FUNCTION "HMI COMMS" : VOID
TITLE =HMI Communications
//OMRON NS12  on DB12
NAME : HMI_COMM
VERSION : 0.1


VAR_TEMP
  UPDATE_PULSE_0 : BOOL ;
  UPDATE_PULSE_1 : BOOL ;
  UPDATE_PULSE_2 : BOOL ;
  UPDATE_PULSE_3 : BOOL ;
  UPDATE_PULSE_4 : BOOL ;
  UPDATE_PULSE_5 : BOOL ;
  UPDATE_PULSE_6 : BOOL ;
  UPDATE_1 : BOOL ;
  UPDATE_2 : BOOL ;
  UPDATE_3 : BOOL ;
  UPDATE_4 : BOOL ;
  UPDATE_5 : BOOL ;
  UPDATE_6 : BOOL ;
  UPDATE_7 : BOOL ;
  UPDATE_8 : BOOL ;
  UPDATE_9 : BOOL ;
  UPDATE_10 : BOOL ;
  UPDATE_11 : BOOL ;
  UPDATE_12 : BOOL ;
  UPDATE_13 : BOOL ;
  TEMP1 : BOOL ;
  TEST : BOOL ;
  CONVEYOR_0_COLOR : BYTE ;
  ELEVATOR_COLOR : BYTE ;
  CONVEYOR_1_COLOR : BYTE ;
  CONVEYOR_2_COLOR : BYTE ;
  CONVEYOR_3_COLOR : BYTE ;
  CONVEYOR_4_COLOR : BYTE ;
  CONVEYOR_5_COLOR : BYTE ;
  CONVEYOR_6_COLOR : BYTE ;
  CONVEYOR_7_COLOR : BYTE ;
  CONVEYOR_8_COLOR : BYTE ;
  CONVEYOR_9_COLOR : BYTE ;
  PUSHER_2_COLOR : BOOL ;
  CONVEYOR_11_COLOR : BYTE ;
  CONVEYOR_12_COLOR : BYTE ;
  CONVEYOR_13_COLOR : BYTE ;
  CONVEYOR_21_COLOR : BYTE ;
  CONVEYOR_22_COLOR : BYTE ;
  CONVEYOR_23_COLOR : BYTE ;
  CONVEYOR_10_COLOR : BYTE ;
  NEW_ORDER_COLOR : BYTE ;
END_VAR
BEGIN
NETWORK
TITLE =HMI - UpDate Timing
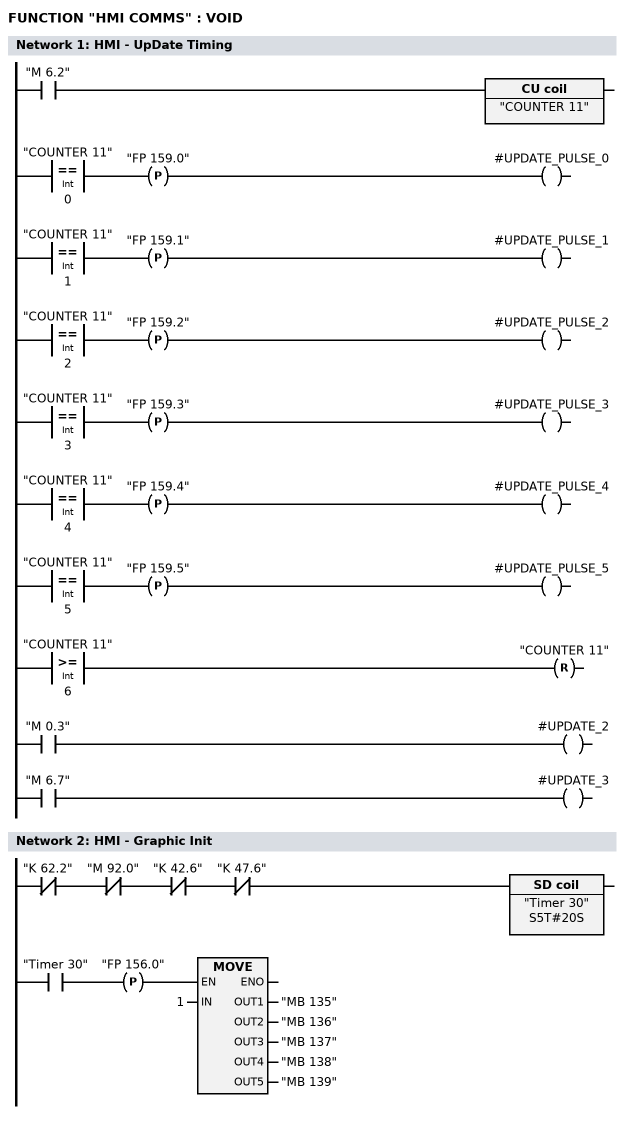

      A     "M 6.2";
      CU    "COUNTER 11";
//;
      A(    ;
      L     "COUNTER 11";
      L     0;
      ==I   ;
      )     ;
      FP    "FP 159.0";
      =     #UPDATE_PULSE_0;
//;
      A(    ;
      L     "COUNTER 11";
      L     1;
      ==I   ;
      )     ;
      FP    "FP 159.1";
      =     #UPDATE_PULSE_1;
//;
      A(    ;
      L     "COUNTER 11";
      L     2;
      ==I   ;
      )     ;
      FP    "FP 159.2";
      =     #UPDATE_PULSE_2;
//;
      A(    ;
      L     "COUNTER 11";
      L     3;
      ==I   ;
      )     ;
      FP    "FP 159.3";
      =     #UPDATE_PULSE_3;
//;
      A(    ;
      L     "COUNTER 11";
      L     4;
      ==I   ;
      )     ;
      FP    "FP 159.4";
      =     #UPDATE_PULSE_4;
//;
      A(    ;
      L     "COUNTER 11";
      L     5;
      ==I   ;
      )     ;
      FP    "FP 159.5";
      =     #UPDATE_PULSE_5;
//;
      A(    ;
      L     "COUNTER 11";
      L     6;
      >=I   ;
      )     ;
      R     "COUNTER 11";
//;;
      A     "M 0.3";
      =     #UPDATE_2;
//;
      A     "M 6.7";
      =     #UPDATE_3;
NETWORK
TITLE =HMI - Graphic Init

      AN    "K 62.2";
      AN    "M 92.0";
      AN    "K 42.6";
      AN    "K 47.6";
      L     S5T#20S;
      SD    "Timer 30";
//;
      A     "Timer 30";
      FP    "FP 156.0";
      JNB   K622;
      L     1;
      T     "MB 135";
      T     "MB 136";
      T     "MB 137";
      T     "MB 138";
      T     "MB 139";

K622: NOP   0;
NETWORK
TITLE =HMI - Doors Monitor

      ON    "E 4.6";
      ON    "E 9.0";
      ON    "E 12.5";
      O     #UPDATE_PULSE_0;
      JNB   DOOR;
      AN    "E 4.6";
      =     "HMI_DB".ELEVATOR_DOOR_STATUS;
//;
      AN    "E 9.0";
      =     "HMI_DB".FLIPPER_DOOR_STATUS;
//;
      AN    "E 12.5";
      =     "HMI_DB".LOADER_DOOR_STATUS;

DOOR: NOP   0;
NETWORK
TITLE =HMI - E-Stop Monitor

      O     "M 1.0";
      O     "M 1.1";
      O     "M 1.2";
      O     "M 1.3";
      O     #UPDATE_PULSE_1;
      JNB   ESTP;
      A     "M 1.0";
      =     "HMI_DB".E_STOP_CONSOLE_STATUS;
//;
      A     "M 1.1";
      =     "HMI_DB".E_STOP_LOADER_STATUS;
//;
      A     "M 1.2";
      =     "HMI_DB".E_STOP_ELEVATOR_STATUS;
//;
      A     "M 1.3";
      =     "HMI_DB".E_STOP_FLIPPER_STATUS;

ESTP: NOP   0;
NETWORK
TITLE =HMI - Motors Fault Status

      A(    ;
      L     "MW 2";
      L     0;
      <>I   ;
      O     ;
      L     "MB 4";
      L     0;
      <>I   ;
      )     ;
      O     "M 7.0";
      O     "M 7.1";
      O     "M 7.2";
      O     #UPDATE_PULSE_2;
      JNB   MTRF;
      A     "M 2.0";
      =     "HMI_DB".CONVEYOR_0_MOTOR_STATUS;
//;
      A     "M 2.1";
      =     "HMI_DB".PUSHER_0_MOTOR_STATUS;
//;
      A     "M 2.2";
      =     "HMI_DB".ELEVATOR_MOTOR_STATUS;
//;
      A     "M 2.3";
      =     "HMI_DB".PUSHER_1_MOTOR_STATUS;
//;
      A     "M 2.4";
      =     "HMI_DB".CONVEYOR_1_MOTOR_STATUS;
//;
      A     "M 2.5";
      =     "HMI_DB".CONVEYOR_2B_MOTOR_STATUS;
//;
      A     "M 2.6";
      =     "HMI_DB".CONVEYOR_2R_MOTOR_STATUS;
//;
      A     "M 2.7";
      =     "HMI_DB".CONVEYOR_3_MOTOR_STATUS;
//;
      A     "M 3.0";
      =     "HMI_DB".CONVEYOR_4_MOTOR_STATUS;
//;
      A     "M 3.1";
      =     "HMI_DB".CONVEYOR_5_MOTOR_STATUS;
//;
      A     "M 3.2";
      =     "HMI_DB".CONVEYOR_6_MOTOR_STATUS;
//;
      A     "M 3.3";
      =     "HMI_DB".CONVEYOR_7_MOTOR_STATUS;
//;
      A     "M 3.4";
      =     "HMI_DB".FLIPPER_MOTOR_STATUS;
//;
      A     "M 3.5";
      =     "HMI_DB".CONVEYOR_8_MOTOR_STATUS;
//;
      A     "M 3.6";
      =     "HMI_DB".TURNTABLE_MOTOR_STATUS;
//;
      A     "M 3.7";
      =     "HMI_DB".CONVEYOR_9_MOTOR_STATUS;
//;
      A     "M 4.0";
      =     "HMI_DB".PUSHER_2_MOTOR_STATUS;
//;
      A     "M 4.1";
      =     "HMI_DB".CONVEYOR_10_MOTOR_STATUS;
//;
      A     "M 4.2";
      =     "HMI_DB".CONVEYOR_11_MOTOR_STATUS;
//;
      A     "M 4.3";
      =     "HMI_DB".CONVEYOR_12_MOTOR_STATUS;
//;
      A     "M 4.4";
      =     "HMI_DB".CONVEYOR_13_MOTOR_STATUS;
//;
      A     "M 4.5";
      =     "HMI_DB".CONVEYOR_21_MOTOR_STATUS;
//;
      A     "M 4.6";
      =     "HMI_DB".CONVEYOR_22_MOTOR_STATUS;
//;
      A     "M 4.7";
      =     "HMI_DB".CONVEYOR_23_MOTOR_STATUS;
//;
      A     "M 7.0";
      =     "HMI_DB".LOADER_LIFT_MOTOR_STATUS;
//;
      A     "M 7.1";
      =     "HMI_DB".LOADER_FING_MOTOR_STATUS;
//;
      A     "M 7.2";
      =     "HMI_DB".LOADER_BELT_MOTOR_STATUS;

MTRF: NOP   0;
NETWORK
TITLE =HMI Light Barriers Status - Conveyors 1, 2, 3 LBs

      A(    ;
      L     IW     5;
      L     "HMI_UPDATE".HMI_GRAPHIC_TOTAL_1;
      <>I   ;
      O     #UPDATE_PULSE_3;
      )     ;
      JNB   LBS1;
      A     "B 5.4";
      =     "HMI_DB".LIGHT_BARRIER_1_STATUS;
//;
      A     "B 5.5";
      =     "HMI_DB".LIGHT_BARRIER_2_STATUS;
//;
      A     "B 6.0";
      =     "HMI_DB".LIGHT_BARRIER_3_STATUS;
//;
      A     "B 6.1";
      =     "HMI_DB".LIGHT_BARRIER_4_STATUS;
//;
      A     "B 6.2";
      =     "HMI_DB".LIGHT_BARRIER_5_STATUS;
//;
      A     "B 6.4";
      =     "HMI_DB".LIGHT_BARRIER_6_STATUS;
//;
      A     "B 5.2";
      =     "HMI_DB".LIGHT_BARRIER_B_STATUS;
//;
      A     "B 5.1";
      =     "HMI_DB".LIGHT_BARRIER_A_STATUS;
//;
      L     IW     5;
      T     "HMI_UPDATE".HMI_GRAPHIC_TOTAL_1;

LBS1: NOP   0;
NETWORK
TITLE =HMI Light Barriers Status - Conveyors 4, 5, 6, 7, 8, 9 LBs

      A(    ;
      L     IW     6;
      L     "HMI_UPDATE".HMI_GRAPHIC_TOTAL_2;
      <>I   ;
      O     #UPDATE_PULSE_4;
      )     ;
      O     "B 8.2";
      JNB   LBS2;
      A     "B 6.7";
      =     "HMI_DB".LIGHT_BARRIER_7_STATUS;
//;
      A     "B 7.0";
      =     "HMI_DB".LIGHT_BARRIER_8_STATUS;
//;
      A     "B 7.1";
      =     "HMI_DB".LIGHT_BARRIER_9_STATUS;
//;
      A     "B 7.2";
      =     "HMI_DB".LIGHT_BARRIER_10_STATUS;
//;
      A     "B 7.3";
      =     "HMI_DB".LIGHT_BARRIER_11_STATUS;
//;
      A     "B 7.4";
      =     "HMI_DB".LIGHT_BARRIER_12_STATUS;
//;
      A     "B 8.2";
      =     "HMI_DB".LIGHT_BARRIER_13_STATUS;
//;
      L     IW     6;
      T     "HMI_UPDATE".HMI_GRAPHIC_TOTAL_2;

LBS2: NOP   0;
NETWORK
TITLE =HMI Light Barriers Status - Conveyors 10, 11, 12, 13, 21, 22, 23

      A(    ;
      L     IW     9;
      L     IW    12;
      +I    ;
      L     IB    15;
      +I    ;
      L     "HMI_UPDATE".HMI_FEED_GRAPHIC;
      <>I   ;
      O     #UPDATE_PULSE_5;
      )     ;
      JNB   LBS3;
      A     "B 9.6";
      =     "HMI_DB".LIGHT_BARRIER_14_STATUS;
//;
      A     "B 9.7";
      =     "HMI_DB".LIGHT_BARRIER_15_STATUS;
//;
      A     "B 10.3";
      =     "HMI_DB".LIGHT_BARRIER_16_STATUS;
//;
      A     "B 10.4";
      =     "HMI_DB".LIGHT_BARRIER_17_STATUS;
//;
      A     "B 10.5";
      =     "HMI_DB".LIGHT_BARRIER_18_STATUS;
//;
      A     "B 10.6";
      =     "HMI_DB".LIGHT_BARRIER_19_STATUS;
//;
      A     "B 10.7";
      =     "HMI_DB".LIGHT_BARRIER_20_STATUS;
//;
      A     "B 11.0";
      =     "HMI_DB".LIGHT_BARRIER_21_STATUS;
//;
      A     "B 11.1";
      =     "HMI_DB".LIGHT_BARRIER_22_STATUS;
//;
      A     "B 11.2";
      =     "HMI_DB".LIGHT_BARRIER_23_STATUS;
//;
      A     "B 12.3";
      =     "HMI_DB".LIGHT_BARRIER_24_STATUS;
//;
      A     "B 13.0";
      =     "HMI_DB".LIGHT_BARRIER_25_STATUS;
//;
      A     "B 15.4";
      =     "HMI_DB".LIGHT_BARRIER_26_STATUS;
//;
      A     "B 15.5";
      =     "HMI_DB".LIGHT_BARRIER_27_STATUS;
//;
      A     "B 15.6";
      =     "HMI_DB".LIGHT_BARRIER_28_STATUS;
//;
      A     "B 15.7";
      =     "HMI_DB".LIGHT_BARRIER_29_STATUS;
//;
      L     IW     9;
      L     IW    12;
      +I    ;
      L     IB    15;
      +I    ;
      T     "HMI_UPDATE".HMI_FEED_GRAPHIC;

LBS3: NOP   0;
NETWORK
TITLE =HMI Light Barriers Status - Conveyors 0 LBs

      A(    ;
      L     QB    62;
      L     "HMI_UPDATE".HMI_MOTOR_TOTAL_1;
      <>I   ;
      O     #UPDATE_PULSE_0;
      )     ;
      O     "B 8.2";
      JNB   LBS4;
      A     "E 34.7";
      =     "HMI_DB".PACKETIZER_GATE_STATUS;
//;
      A     "B 35.2";
      =     "HMI_DB".LIGHT_BARRIER_30_STATUS;
//;
      A     "B 35.3";
      =     "HMI_DB".LIGHT_BARRIER_31_STATUS;
//;
      A     "B 35.4";
      =     "HMI_DB".LIGHT_BARRIER_32_STATUS;
//;
      L     QB    62;
      T     "HMI_UPDATE".HMI_MOTOR_TOTAL_1;

LBS4: NOP   0;
NETWORK
TITLE =HMI Prox Sensors Status - Elevator - Proxs

      A(    ;
      L     IB     4;
      L     "HMI_UPDATE".HMI_ELEVATOR_PROXS;
      <>I   ;
      O     #UPDATE_PULSE_1;
      )     ;
      JNB   PRX1;
      AN    "P 4.0";
      =     "HMI_DB".PROX_1_STATUS;
//;
      AN    "P 4.1";
      =     "HMI_DB".PROX_2_STATUS;
//;
      AN    "P 4.2";
      =     "HMI_DB".PROX_3_STATUS;
//;
      AN    "P 4.3";
      =     "HMI_DB".PROX_4_STATUS;
//;
      AN    "P 4.4";
      =     "HMI_DB".PROX_5_STATUS;
//;
      AN    "P 4.5";
      =     "HMI_DB".PROX_6_STATUS;
//;
      L     IB     4;
      T     "HMI_UPDATE".HMI_ELEVATOR_PROXS;

PRX1: NOP   0;
NETWORK
TITLE =HMI Prox Sensors Status - Flipper / TurnTable - Proxs

      A(    ;
      L     IW     8;
      L     "HMI_UPDATE".HMI_FLIPPER_PROXS;
      <>I   ;
      O     #UPDATE_PULSE_2;
      )     ;
      JNB   PRX2;
      AN    "P 8.0";
      =     "HMI_DB".PROX_8_STATUS;
//;
      AN    "P 8.1";
      =     "HMI_DB".PROX_7_STATUS;
//;
      AN    "P 8.5";
      =     "HMI_DB".PROX_9_STATUS;
//;
      AN    "P 8.6";
      =     "HMI_DB".PROX_10_STATUS;
//;
      AN    "P 9.2";
      =     "HMI_DB".PROX_11_STATUS;
//;
      AN    "P 9.3";
      =     "HMI_DB".PROX_12_STATUS;
//;
      L     IW     8;
      T     "HMI_UPDATE".HMI_FLIPPER_PROXS;

PRX2: NOP   0;
NETWORK
TITLE =HMI Prox Sensors Status - Pusher 2 / Pivot 10 - Proxs

      A(    ;
      L     IB    10;
      L     IB    15;
      +I    ;
      L     "HMI_UPDATE".HMI_PUSHER_PROXS;
      <>I   ;
      O     #UPDATE_PULSE_3;
      )     ;
      JNB   PRX3;
      AN    "P 10.0";
      =     "HMI_DB".PROX_13_STATUS;
//;
      AN    "P 10.1";
      =     "HMI_DB".PROX_14_STATUS;
//;
      A     "P 15.0";
      =     "HMI_DB".PROX_15_STATUS;
//;
      A     "P 15.1";
      =     "HMI_DB".PROX_16_STATUS;
//;
      L     IB    10;
      L     IB    15;
      +I    ;
      T     "HMI_UPDATE".HMI_PUSHER_PROXS;

PRX3: NOP   0;
NETWORK
TITLE =HMI Prox Sensors Status - Feeder - Proxs

      A(    ;
      L     IW    11;
      L     IB    13;
      +I    ;
      L     "HMI_UPDATE".HMI_FEEDER_PROXS;
      <>I   ;
      O     #UPDATE_PULSE_4;
      )     ;
      JNB   PRX4;
      AN    "P 13.2";
      =     "HMI_DB".PROX_17_STATUS;
//;
      AN    "P 13.1";
      =     "HMI_DB".PROX_18_STATUS;
//;
      AN    "P 11.4";
      =     "HMI_DB".PROX_19_STATUS;
//;
      AN    "P 11.5";
      =     "HMI_DB".PROX_20_STATUS;
//;
      AN    "P 11.6";
      =     "HMI_DB".PROX_21_STATUS;
//;
      AN    "P 11.7";
      =     "HMI_DB".PROX_22_STATUS;
//;
      A     "P 12.0";
      =     "HMI_DB".PROX_23_STATUS;
//;
      A     "P 12.1";
      =     "HMI_DB".PROX_24_STATUS;
//;
      L     IW    11;
      L     IB    13;
      +I    ;
      T     "HMI_UPDATE".HMI_FEEDER_PROXS;

PRX4: NOP   0;
NETWORK
TITLE =HMI - Pusher 0 - Graphic

      A(    ;
      O     "K 62.2";
      O     "K 62.3";
      O     #UPDATE_PULSE_5;
      )     ;
      JNB   PUS0;
      A     "K 62.2";
      AN    "K 62.3";
      A     "M 6.1";
      AN(   ;
      L     "MB 135";
      L     L#128;
      >=I   ;
      )     ;
      FP    "FP 156.1";
      JNB   E622;
      L     "MB 135";
      SLW   1;
      T     "MB 135";

E622: NOP   0;

      A     "K 62.3";
      AN    "K 62.2";
      A     "M 6.1";
      AN(   ;
      L     "MB 135";
      L     L#1;
      <=I   ;
      )     ;
      FP    "FP 156.2";
      JNB   R623;
      L     "MB 135";
      SRW   1;
      T     "MB 135";

R623: NOP   0;

      A     "M 6.1";
      FP    "HMI_DB".FP133;
      JNB   P133;
      L     L#255;
      L     "MB 135";
      -I    ;
      T     DB12.DBB    4;

P133: NOP   0;

PUS0: NOP   0;
NETWORK
TITLE =HMI - Elevator - Graphic

      A(    ;
      O     "M 92.0";
      O     "M 92.1";
      O     #UPDATE_PULSE_0;
      )     ;
      JNB   ELEV;
      A     "M 92.0";
      AN    "M 92.1";
      A     "M 6.2";
      AN(   ;
      L     "MB 136";
      L     L#128;
      >=I   ;
      )     ;
      FP    "FP 156.3";
      JNB   R420;
      L     "MB 136";
      SLW   1;
      T     "MB 136";

R420: NOP   0;

      A     "M 92.1";
      AN    "M 92.0";
      A     "M 6.2";
      AN(   ;
      L     "MB 136";
      L     L#1;
      <=I   ;
      )     ;
      FP    "FP 156.4";
      JNB   F420;
      L     "MB 136";
      SRW   1;
      T     "MB 136";

F420: NOP   0;

      A     "M 6.2";
      FP    "HMI_DB".FP134;
      JNB   P134;
      L     L#255;
      L     "MB 136";
      -I    ;
      T     DB12.DBB    5;

P134: NOP   0;

ELEV: NOP   0;
NETWORK
TITLE =HMI - Pusher 1 - Graphic

      A(    ;
      O     "K 42.6";
      O     "K 42.7";
      O     #UPDATE_PULSE_1;
      )     ;
      JNB   PUS1;
      A     "K 42.6";
      AN    "K 42.7";
      A     "M 6.1";
      AN(   ;
      L     "MB 137";
      L     L#128;
      >=I   ;
      )     ;
      FP    "FP 156.5";
      JNB   E426;
      L     "MB 137";
      SLW   1;
      T     "MB 137";

E426: NOP   0;

      A     "K 42.7";
      AN    "K 42.6";
      A     "M 6.1";
      AN(   ;
      L     "MB 137";
      L     L#1;
      <=I   ;
      )     ;
      FP    "FP 156.6";
      JNB   R427;
      L     "MB 137";
      SRW   1;
      T     "MB 137";

R427: NOP   0;

      A     "M 6.1";
      FP    "HMI_DB".FP135;
      JNB   P135;
      L     L#255;
      L     "MB 137";
      -I    ;
      T     DB12.DBB    6;

P135: NOP   0;

PUS1: NOP   0;
NETWORK
TITLE =HMI - Flipper Graphic

      A(    ;
      O     "K 46.0";
      O     "K 46.1";
      O     #UPDATE_PULSE_2;
      )     ;
      JNB   FLPN;
      L     3;
      A     "P 8.0";
      A     "P 8.1";
      JC    FLIP;
      L     0;

FLIP: T     "HMI_DB".FLIPPER_TURN_COLOR;

      L     1;
      AN    "P 8.0";
      A     "P 8.1";
      JC    CCW1;
      L     "HMI_DB".FLIPPER_TURN_COLOR;

CCW1: T     "HMI_DB".FLIPPER_CCW;

      L     1;
      AN    "P 8.1";
      A     "P 8.0";
      JC    CW1;
      L     "HMI_DB".FLIPPER_TURN_COLOR;

CW1:  T     "HMI_DB".FLIPPER_CW;

      L     6;
      A     "M 42.0";
      JC    FLON;
      L     9;

FLON: T     "HMI_DB".FLIPPER_COLOR;

FLPN: NOP   0;
NETWORK
TITLE =HMI - TurnTable Graphic

      A(    ;
      O     "A 47.0";
      O     "A 47.1";
      O     #UPDATE_PULSE_3;
      )     ;
      JNB   TURN;
      A(    ;
      ON    "P 9.2";
      ON    "P 9.3";
      )     ;
      S     "HMI_DB".TURNTABLE_DELIV_POSITION;
//;
      A(    ;
      ON    "P 8.5";
      ON    "P 8.6";
      )     ;
      R     "HMI_DB".TURNTABLE_DELIV_POSITION;
//;
      AN    "M 7.3";
      =     "HMI_DB".TURNTABLE_REVERSE_ARROW;
//;
      A     "M 7.3";
      =     "HMI_DB".TURNTABLE_DIR_SELECT_SW;

TURN: NOP   0;

NETWORK
TITLE =HMI - Pusher 2 - Graphic

      A(    ;
      O     "K 47.6";
      O     "K 47.7";
      O     #UPDATE_PULSE_4;
      )     ;
      JNB   PUS2;
      A     "K 47.6";
      AN    "K 47.7";
      A     "M 6.1";
      AN(   ;
      L     "MB 138";
      L     L#128;
      >=I   ;
      )     ;
      FP    "FP 156.7";
      JNB   E476;
      L     "MB 138";
      SLW   1;
      T     "MB 138";

E476: NOP   0;

      A     "K 47.7";
      AN    "K 47.6";
      A     "M 6.1";
      AN(   ;
      L     "MB 138";
      L     L#1;
      <=I   ;
      )     ;
      FP    "FP 157.0";
      JNB   R477;
      L     "MB 138";
      SRW   1;
      T     "MB 138";

R477: NOP   0;

      A     "M 6.1";
      FP    "HMI_DB".FP140;
      JNB   P140;
      L     L#255;
      L     "MB 138";
      -I    ;
      T     DB12.DBB    7;

P140: NOP   0;

PUS2: NOP   0;
NETWORK
TITLE =HMI - Pivot Graphic

      A(    ;
      O     "K 53.0";
      O     "K 53.1";
      O     #UPDATE_PULSE_5;
      )     ;
      JNB   PIVO;
      AN    "P 15.1";
      =     DB12.DBX   88.1;
//;
      AN    "P 15.0";
      =     DB12.DBX   88.0;
//;
      AN    "P 15.0";
      AN    "P 15.1";
      =     DB12.DBX   88.2;

PIVO: NOP   0;
NETWORK
TITLE =HMI - Feeder Graphic

      A(    ;
      L     IW    11;
      L     IB    13;
      +I    ;
      L     "HMI_UPDATE".HMI_FEEDER_GRAPHIC;
      <>I   ;
      O     #UPDATE_PULSE_0;
      )     ;
      JNB   FEED;

      A     "P 13.2";
      AN    "P 11.4";
      O     ;
      A     "P 11.5";
      AN    "P 11.4";
      JNB   M131;
      L     L#64;
      T     "MB 139";

M131: NOP   0;

      AN    "P 13.2";
      AN    "P 13.1";
      AN    "P 11.4";
      JNB   M132;
      L     L#128;
      T     "MB 139";

M132: NOP   0;

      AN    "P 11.4";
      AN    "P 11.5";
      JNB   M114;
      L     L#32;
      T     "MB 139";

M114: NOP   0;

      A     "P 11.4";
      AN    "P 11.5";
      A     "A 50.1";
      S     "M 70.5";
//;
      A(    ;
      A     "M 70.6";
      A     "A 50.0";
      AN    "P 11.5";
      O     ;
      A     "M 70.5";
      A     "A 50.1";
      )     ;
      JNB   M115;
      L     L#16;
      T     "MB 139";
      R     "M 70.6";

M115: NOP   0;

      A     "P 11.7";
      AN    "P 11.6";
      A     "A 50.0";
      S     "M 70.6";
//;
      A(    ;
      A     "M 70.5";
      A     "A 50.1";
      AN    "P 11.6";
      O     ;
      A     "M 70.6";
      A     "A 50.0";
      )     ;
      JNB   M116;
      L     L#8;
      T     "MB 139";
      R     "M 70.5";

M116: NOP   0;

      AN    "E 12.2";
      AN    "P 11.7";
      AN    "P 12.1";
      JNB   M117;
      L     L#4;
      T     "MB 139";

M117: NOP   0;

      AN    "E 12.2";
      AN    "P 11.7";
      A     "P 12.1";
      JNB   M121;
      L     L#6;
      T     "MB 139";

M121: NOP   0;

      A     "E 12.2";
      AN    "P 11.7";
      A     "P 12.1";
      JNB   M122;
      L     L#1;
      T     "MB 139";

M122: NOP   0;

      A     "M 6.2";
      FP    "HMI_DB".FP141;
      JNB   P141;
      L     L#255;
      L     "MB 139";
      -I    ;
      T     DB12.DBB   19;

P141: NOP   0;

      L     IW    11;
      L     IB    13;
      +I    ;
      T     "HMI_UPDATE".HMI_FEEDER_GRAPHIC;

FEED: NOP   0;
NETWORK
TITLE =HMI - Motor Run Status

      A(    ;
      L     QW    42;
      L     QW    44;
      +I    ;
      L     QW    46;
      +I    ;
      L     QW    48;
      +I    ;
      L     QW    50;
      +I    ;
      L     QB    53;
      +I    ;
      L     QB    54;
      +I    ;
      L     "HMI_UPDATE".HMI_MOTOR_GRAPHIC;
      <>I   ;
      O     #UPDATE_PULSE_1;
      )     ;
      JNB   MTR;
      O     "K 62.0";
      O     "K 62.1";
      L     0;
      JCN   K620;
      A     "K 62.0";
      L     3;
      JC    K620;
      L     6;
K620: T     "HMI_DB".CONV_0_COLOR_WORD;

      L     5;
      A     "M 14.7";
      O     "M 100.2";
      JC    E00;
      L     0;
E00:  T     #ELEVATOR_COLOR;

      L     #ELEVATOR_COLOR;
      O     "M 92.0";
      O     "M 92.1";
      JCN   Q420;
      A     "M 92.0";
      L     3;
      JC    Q420;
      L     6;
Q420: T     "HMI_DB".ELEVATOR_COLOR_WORD;

      L     0;
      A(    ;
      O     "K 42.6";
      O     "K 42.7";
      )     ;
      JCN   Q427;
      L     3;
Q427: T     "HMI_DB".PUSHER_1_COLOR_WORD;

      L     0;
      A     "A 43.0";
      JCN   Q430;
      L     3;
Q430: T     "HMI_DB".CONV_1_COLOR_WORD;

      L     5;
      A     "M 22.7";
      O     "M 100.5";
      JC    C02;
      L     0;
C02:  T     #CONVEYOR_2_COLOR;

      L     #CONVEYOR_2_COLOR;
      A     "K 43.4";
      JCN   Q434;
      L     3;
Q434: T     "HMI_DB".CONV_2_BELT_COLOR_WORD;

      L     0;
      A     "Y 43.6";
      JCN   Q436;
      L     3;
Q436: T     "HMI_DB".LIFT_ROLLER_2_COLOR_WORD;

      L     0;
      A     "K 43.5";
      JCN   Q435;
      L     3;
Q435: T     "HMI_DB".CONV_2_ROLLER_COLOR_WORD;

      L     0;
      A     "A 44.0";
      JCN   Q440;
      L     3;
Q440: T     "HMI_DB".CONV_3_COLOR_WORD;

      L     5;
      A     "M 30.7";
      O     "M 102.0";
      JC    C04;
      L     0;
C04:  T     #CONVEYOR_4_COLOR;

      L     #CONVEYOR_4_COLOR;
      A     "A 44.3";
      AN    "M 31.5";
      JCN   Q443;
      L     6;
Q443: T     "HMI_DB".CONV_4_COLOR_WORD;

      A     "A 44.3";
      A     "M 31.5";
      JNB   M315;
      L     3;
      T     "HMI_DB".CONV_4_COLOR_WORD;

M315: NOP   0;

      L     0;
      A     "A 45.0";
      JCN   Q450;
      L     3;
Q450: T     "HMI_DB".CONV_5_COLOR_WORD;

      L     5;
      A     "M 38.7";
      O     "M 102.2";
      JC    C06;
      L     0;
C06:  T     #CONVEYOR_6_COLOR;

      L     #CONVEYOR_6_COLOR;
      A     "A 45.3";
      JCN   Q453;
      L     3;
Q453: T     "HMI_DB".CONV_6_COLOR_WORD;

      L     5;
      A     "M 42.7";
      O     "M 102.3";
      JC    C07;
      L     0;
C07:  T     #CONVEYOR_7_COLOR;

      L     #CONVEYOR_7_COLOR;
      A     "A 45.6";
      JCN   Q456;
      L     3;
Q456: T     "HMI_DB".CONV_7_COLOR_WORD;

      L     0;
      A(    ;
      O     "K 46.0";
      O     "K 46.1";
      )     ;
      JCN   Q461;
      L     3;
Q461: T     "HMI_DB".FLIPPER_COLOR_WORD;

      L     0;
      A(    ;
      O     "A 47.0";
      O     "A 47.1";
      )     ;
      JCN   A470;
      L     7;

A470: T     "HMI_DB".TURN_COLOR;

//      L     0
//      AN    "M 6.2"
//      A(
//      O     "A 47.0"
//      O     "A 47.1"
//      )
//      JCN   A471
//      L     7

//A471: T     "HMI_DB".HMI_TURN_COLOR

      L     "HMI_DB".TURN_COLOR;
      A(    ;
      O     "A 46.4";
      O     "A 46.5";
      )     ;
      JCN   Q464;
      L     3;
Q464: T     "HMI_DB".CONV_8_COLOR_WORD;

      L     0;
      A     "A 47.0";
      JCN   Q470;
      L     3;
Q470: T     "HMI_DB".TURN_TABLE_COLOR_WORD;

      L     0;
      A     "K 47.5";
      JCN   Q475;
      L     3;
Q475: T     "HMI_DB".CONV_9_COLOR_WORD;

      L     0;
      A(    ;
      O     "K 47.6";
      O     "K 47.7";
      )     ;
      JCN   Q477;
      L     3;
Q477: T     "HMI_DB".PUSHER_2_COLOR_WORD;

      L     5;
      A     "M 98.1";
      O     "M 98.2";
      O     "M 106.1";
      JC    C10;
//;
      L     4;
      A     "M 55.4";
      A     "M 8.4";
      A     "M 6.5";
      JC    C10;
      L     0;

C10:  T     #CONVEYOR_10_COLOR;

      L     #CONVEYOR_10_COLOR;
      A     "A 48.0";
      A(    ;
      ON    "M 55.5";
      ON    "M 10.0";
      )     ;
      JCN   Q480;
      L     6;
Q480: T     "HMI_DB".CONV_10_COLOR_WORD;

      A     "A 48.0";
      A(    ;
      O     "M 55.5";
      O     "M 10.0";
      )     ;
      JNB   M555;
      L     3;
      T     "HMI_DB".CONV_10_COLOR_WORD;

M555: NOP   0;


      L     0;
      A     "A 48.3";
      JCN   Q483;
      L     3;
Q483: T     "HMI_DB".CONV_11_COLOR_WORD;

      L     0;
      A     "A 48.6";
      JCN   Q486;
      L     3;
Q486: T     "HMI_DB".CONV_12_COLOR_WORD;

      L     5;
      A     "M 66.7";
      O     "M 106.4";
      JC    C13;
      L     0;
C13:  T     #CONVEYOR_13_COLOR;

      L     #CONVEYOR_13_COLOR;
      A     "A 49.0";
      JCN   Q490;
      L     3;
Q490: T     "HMI_DB".CONV_13_COLOR_WORD;

      L     0;
      A     "A 53.4";
      JCN   Q534;
      L     3;
Q534: T     "HMI_DB".CONV_21_COLOR_WORD;

      L     0;
      A     "A 53.6";
      JCN   Q536;
      L     3;
Q536: T     "HMI_DB".CONV_22_COLOR_WORD;

      L     5;
      A     "M 86.7";
      O     "M 106.7";
      JC    C23;
      L     0;
C23:  T     #CONVEYOR_23_COLOR;

      L     #CONVEYOR_23_COLOR;
      A     "A 54.0";
      JCN   Q540;
      L     3;
Q540: T     "HMI_DB".CONV_23_COLOR_WORD;

      A     "M 0.7";
      =     "HMI_DB".COMPRESSED_AIR;
//;
      O     "A 50.0";
      O     "A 50.1";
      L     0;
      JCN   Q500;
      A     "A 50.0";
      L     3;
      JC    Q500;
      L     6;
Q500: T     "HMI_DB".LOADER_LIFT_COLOR_WORD;

      L     0;
      A     "A 51.0";
      JCN   Q510;
      L     3;
Q510: T     "HMI_DB".FINGERS_BELT_COLOR_WORD;

      L     QW    42;
      L     QW    44;
      +I    ;
      L     QW    46;
      +I    ;
      L     QW    48;
      +I    ;
      L     QW    50;
      +I    ;
      L     QB    53;
      +I    ;
      L     QB    54;
      +I    ;
      T     "HMI_UPDATE".HMI_MOTOR_GRAPHIC;

MTR:  NOP   0;
END_FUNCTION

